Fanuc KAREL source: kb00162.KL

PROGRAM KB00162
%NOLOCKGROUP
VAR
P1:INTEGER;P2:INTEGER;P3 : XYZWPREXT;P4:INTEGER
BEGIN
--
--
--
P1=1
P2=1
P4=1
SET_EPOS_TPE(P1,P2,P3,P4,1)
END KB00162
